Fanuc KAREL source: KD00041.KL

PROGRAM KD00041
%NOLOCKGROUP
%ENVIRONMENT UIF
VAR
  I: INTEGER
  J: INTEGER
  B: BOOLEAN
  R: REAL
  S: STRING[80]
  D: DISP_DAT_T
BEGIN
  I = 1
END KD00041
